{attribute 'linkalways'} 
{attribute 'no_explicit_call' := 'This FB is a CLASS and must be accessed using methods or properties'}
{attribute 'enable_dynamic_creation'}
FUNCTION_BLOCK _Array0to1OfDINT EXTENDS ArrayDatatypeBase_1D
VAR CONSTANT
	lBound : DINT := 0;
	uBound : DINT := 1;
END_VAR
VAR
	localData : ARRAY [lBound..uBound] OF DINT;
	activeData : REFERENCE TO ARRAY [lBound..uBound] OF DINT REF= localData;
	elements : ARRAY [lBound..uBound] OF _DINT(0);
	baseType : _DINT(0);
END_VAR

PROPERTY PUBLIC Address : PVOID
GET
Address := ADR(activeData);
END_GET
END_PROPERTY

PROPERTY PUBLIC BaseDatatype : I_Datatype
GET
BaseDatatype := baseType;
END_GET
END_PROPERTY

METHOD PUBLIC ClearReference
VAR_INPUT
END_VAR
activeData REF= localData;
SetElementReference();
END_METHOD

METHOD PUBLIC Clone : I_Datatype
VAR
    pClone : POINTER TO _Array0to1OfDINT;
END_VAR
pClone := __NEW(_Array0to1OfDINT());
pClone^.Value := Value;
Clone := pClone^;
END_METHOD

METHOD FB_init : BOOL
VAR_INPUT
	bInitRetains : BOOL; // if TRUE, the retain variables are initialized (warm start / cold start)
	bInCopyCode : BOOL;  // if TRUE, the instance afterwards gets moved into the copy code (online change)
END_VAR
SetElementReference();
END_METHOD

METHOD PUBLIC MakeReferenceTo
VAR_INPUT
	ReferenceTarget : REFERENCE TO ARRAY [lBound..uBound] OF DINT;
END_VAR
activeData REF= ReferenceTarget;
SetElementReference();
END_METHOD

METHOD PROTECTED OnSerializeArrayValues
VAR_INPUT
	Serializer : I_Serializer;
END_VAR
VAR
	i : DINT;
END_VAR
FOR i := lBound TO uBound DO
	elements[i].SerializeWith(Serializer);
END_FOR
END_METHOD

METHOD PROTECTED SetElementReference
VAR_INPUT
END_VAR
VAR
	i : DINT;
END_VAR
FOR i := lBound TO uBound DO
	elements[i].MakeReferenceTo(activeData[i]);
END_FOR
END_METHOD

PROPERTY PUBLIC Size : UDINT
GET
Size := SIZEOF(activeData);
END_GET
END_PROPERTY

METHOD PROTECTED TryDeserializeArrayValues : BOOL
VAR_INPUT
	Deserializer : I_Deserializer;
	Feedback : I_DeserializerFeedback;
END_VAR
VAR
	failed : BOOL;
	enumerator : I_DeserializerArrayForwardEnumerator;
	i : DINT;
END_VAR
enumerator := Deserializer.GetArrayEnumerator();
i := lBound;

WHILE enumerator.MoveNext() AND i <= uBound AND NOT failed DO
	
	IF NOT elements[i].TryDeserializeFrom(enumerator.Current, Feedback) THEN
		failed := TRUE;
		EXIT;
	END_IF
	i := i + 1;

END_WHILE
enumerator.Dispose();

TryDeserializeArrayValues := NOT failed;
END_METHOD

METHOD PUBLIC TryGetElementAsDatatypeByIndex : BOOL
VAR_INPUT
	Index : DINT;
	Destination : REFERENCE TO I_Datatype;
END_VAR
IF Index < lbound OR Index > ubound THEN
	RETURN;
END_IF

Destination := elements[Index];
TryGetElementAsDatatypeByIndex := TRUE;
END_METHOD

METHOD PUBLIC TryGetLowerBound : BOOL
VAR_INPUT
	Dimention : UDINT;
	Destination : REFERENCE TO DINT;
END_VAR
IF Dimention = 1 THEN
	Destination := lBound;
	TryGetLowerBound := TRUE;
END_IF
END_METHOD

METHOD PUBLIC TryGetUpperBound : BOOL
VAR_INPUT
	Dimention : UDINT;
	Destination : REFERENCE TO DINT;
END_VAR
IF Dimention = 1 THEN
	Destination := uBound;
	TryGetUpperBound := TRUE;
END_IF
END_METHOD

METHOD TryMakeReferenceTo : BOOL
VAR_INPUT
	Target : I_Datatype;
END_VAR
VAR
	pTargetData : POINTER TO ARRAY [lBound..uBound] OF DINT;
END_VAR
IF NOT IsEquivalentTo(Target) THEN
	RETURN;
END_IF

pTargetData := Target.Address;
activeData REF= pTargetData^;
SetElementReference();
TryMakeReferenceTo := TRUE;
END_METHOD

PROPERTY PUBLIC Value : REFERENCE TO ARRAY [lBound..uBound] OF DINT;
GET
Value ref= activeData;
END_GET
END_PROPERTY

END_FUNCTION_BLOCK

(* stored: Version 1.1.0.1, ProductVersion 3.1.4024.13
   POU _Array0to1OfDINT: Id {04116934-13ab-050b-00a4-03ef308ac515}, SpecialFunc None
   Folder Core: Id {d74209f3-d5cb-0df4-1aad-bc6d2dcb6ddd}
   Folder Constructor: Id {d042b0d5-847b-0f80-0768-6e4a99292f78}
   Folder Protected: Id {19fdcc57-cf51-01d1-2a0b-0a75cbd9a149}
   Folder Customize: Id {88ba6ca0-79b6-0ac6-29e3-a1b90c09d5f4}
   Property Address: Id {d3a5bef2-5cb6-0652-18e2-60a3ccfe31d2}
   Get Get: Id {e73cac45-e663-0545-2cc0-414d1d0311e1}
   Property BaseDatatype: Id {0269d541-bad7-0d9a-0e4c-bdd91210c592}
   Get Get: Id {95dfb333-a2e6-02ad-00bf-e64d2c71d51c}
   Method ClearReference: Id {faaabd2e-4e48-08ee-0037-ee73915006fd}
   Method Clone: Id {a692bc0a-278c-0046-0f76-ebd148cffd6a}
   Method FB_init: Id {7df8f189-d944-0ddf-368b-f072c70a0398}
   Method MakeReferenceTo: Id {9e27c148-ad2b-0b65-2d7f-ab4071d38e42}
   Method OnSerializeArrayValues: Id {c139ab03-e366-0f77-3b68-e8484efc0829}
   Method SetElementReference: Id {59b59883-1d59-039b-05f6-6094f0d97e04}
   Property Size: Id {16d5768d-c229-02a1-2ae1-99320dd01e12}
   Get Get: Id {9111c6bd-1ccf-01ba-2027-cad2a3541567}
   Method TryDeserializeArrayValues: Id {3f5d950c-0e85-00f5-3e2d-60dba720e040}
   Method TryGetElementAsDatatypeByIndex: Id {8319e015-e240-0a1c-307a-44932d2e484d}
   Method TryGetLowerBound: Id {ebd7953d-4142-02f9-2d18-981ef043c927}
   Method TryGetUpperBound: Id {9c9de581-e1ae-0ea5-0f01-7f2047f16e23}
   Method TryMakeReferenceTo: Id {29e53d4d-535b-01ea-0307-6ce40a60fa38}
   Property Value: Id {2ce8155d-7f66-06b6-3502-2baee3f8f8eb}
   Get Get: Id {761f0404-c759-05a2-2618-3c3cd8beb2d7} *)
